(*
Section Title
-------------
This document consists of two main sections and several subsections. All text blocks up to the next title of the same or higher level
are included in a section (or subsection, etc.).

================
1. Section Title
================
Sections are identified through their titles, which are marked up with adornment:
"underlines" below the title text, or underlines and matching "overlines" above the title.

-----------------
1.1 Section Title
-----------------
A document must be consistent in its use of section titles: once a hierarchy of title styles is established,
sections must use that hierarchy.
Rather than imposing a fixed number and order of section title adornment styles,
the order enforced will be the order as encountered.
The first style encountered will be an outermost title, the second style will be a subtitle,
the third will be a subsubtitle, and so on.

1.2.1 Section Title
===================
Underline-only adornment styles are distinct
from overline-and-underline styles that use the same character. 

1.2.1.1 Section Title
*********************
An underline/overline is a single repeated punctuation character that begins in column 1
and forms a line extending at least as far as the right edge of the title text.

1.2.1.2 Section Title
*********************

1.2.2 Section Title
===================

-----------------
1.2 Section Title
-----------------

=================
2. Section Title
=================

-----------------
2.1 Section Title
-----------------
*)

FUNCTION_BLOCK FB_Libdoc_Sections
VAR_INPUT
    nVarA : INT;
    nVarB : INT;
END_VAR
VAR_OUTPUT
    nSum : INT;
END_VAR
VAR
END_VAR

END_FUNCTION_BLOCK

(* stored: Version 1.1.0.1, ProductVersion 3.1.4022.17
   POU FB_Libdoc_Sections: Id {892b6f99-49d7-4a88-8149-92f13a5881b1}, SpecialFunc None *)
